FUNCTION_BLOCK FsServer (* Status and messages of the own file server of logiBUS *)
  (* Standard: 61499-2; Description: The own ISO 11783-13 file server of logiBUS: one volume \\LOGIBUS\ = /data/fs with quota. \n Switched on with PART_13_FS = 1 in /data/functionalities.ini (restart), quota PART_13_FS_QUOTA_KB, bus share PART_13_FS_BUS_SHARE. \n IND for every file a client has written (closed after writing), with the local path. \n CHG when bRunning, u8Clients or u8OpenFiles changes (no polling with REQ needed). \n Only one FsServer per device: a second instance takes the messages over. *)
  (* Version 1.0, 2026-11-26, Franz Höpfinger, initial API and implementation and/or initial documentation *)
  PACKAGE isobus::fs_server;
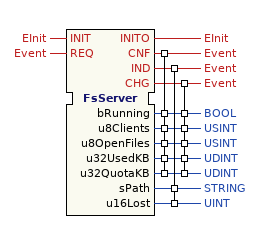
  EVENT_INPUT
    INIT : EInit; (* Service Initialization *)
    REQ; (* Read the status *)
  END_EVENT
  EVENT_OUTPUT
    INITO : EInit; (* Initialization Confirm *)
    CNF WITH bRunning, u8Clients, u8OpenFiles, u32UsedKB, u32QuotaKB; (* Status read *)
    IND WITH sPath, u16Lost; (* A client has written a file *)
    CHG WITH bRunning, u8Clients, u8OpenFiles, u32UsedKB, u32QuotaKB; (* Status changed (running, clients, open files) *)
  END_EVENT
  VAR_OUTPUT
    bRunning : BOOL; (* Server switched on and address claimed *)
    u8Clients : USINT; (* Connected clients *)
    u8OpenFiles : USINT; (* Open files of all clients *)
    u32UsedKB : UDINT; (* Bytes below /data/fs in KB (updated every 10 s) *)
    u32QuotaKB : UDINT; (* Quota of /data/fs in KB *)
    sPath : STRING; (* With IND: local path of the written file, e.g. /data/fs/IMPORT/a.xml *)
    u16Lost : UINT; (* With IND: messages lost before this one (queue of 16 full) *)
  END_VAR
END_FUNCTION_BLOCK
